(* IEC 61131-3 sources: plcassist-cli/packages/volt-lsp-iec/test-corpus/pro2193/Device/Plc Logic/Application/09 Misc, 1 file *)

(* ---- GVL_Exceptions.gvl ---- *)
{attribute 'qualified_only'}
VAR_GLOBAL
	xException : BOOL;
	aeExceptionCodes: ARRAY[0..50] OF __SYSTEM.ExceptionCode;
	iCounter	: UDINT;
END_VAR
